(* Error Buzzer Blinky *)

PROGRAM main
  VAR
    FaultActive AT %MX0.0 : BOOL; (* Input Variable *)
    Buzzer AT %QX0.2 : BOOL;
    TON0 : TON;
    TOF0 : TOF;
  END_VAR

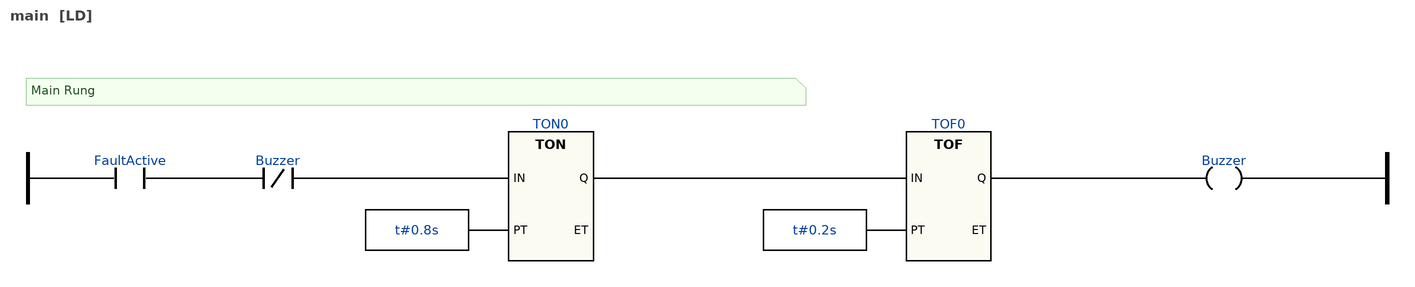
(* LD diagram, written out as Structured Text *)
(* Main Rung *)
TON0(IN := FaultActive AND NOT Buzzer, PT := t#0.8s);
TOF0(IN := TON0.Q, PT := t#0.2s);
Buzzer := TOF0.Q;
END_PROGRAM
